Fanuc KAREL source: kd00015.KL

-- PROVISIONAL review KL for V770-1; original PC SHA256 4509d865207344b37e3f2777ffe3726d0b491e45a606fccd107e2c295447d1f1
-- Incomplete behavior may be omitted. Consult companion uncertainty JSON. Do not deploy.
PROGRAM KD00015
%NOLOCKGROUP
VAR
  I : INTEGER
  J : INTEGER
  B : BOOLEAN
  R : REAL
  S : STRING[80]
BEGIN
  -- UNRESOLVED_PC offsets 5-6; opcodes 16
  -- UNRESOLVED_PC offsets 11-15; opcodes 7F
END KD00015
